// TIA Portal V20 export
Screen "CycleTime"  1276x673
  ScreenItem "Faceplate container_1" at 135,81 size 64x420  Type=HmiFaceplateContainer
  ScreenItem "Line_22" at 128,84 size 1x400  Type=HmiLine
  ScreenItem "Line_46" at 110,355 size 17x0  Type=HmiLine
  ScreenItem "Line_47" at 111,420 size 17x0  Type=HmiLine
  ScreenItem "Line_48" at 112,484 size 17x0  Type=HmiLine
  ScreenItem "Casella di testo_56" at 62,271 size 48x30  Type=HmiTextBox
  ScreenItem "Casella di testo_57" at 62,339 size 48x30  Type=HmiTextBox
  ScreenItem "Casella di testo_59" at 62,405 size 48x30  Type=HmiTextBox
  ScreenItem "Casella di testo_60" at 62,468 size 48x30  Type=HmiTextBox
  ScreenItem "Line_49" at 109,224 size 17x0  Type=HmiLine
  ScreenItem "Casella di testo_7" at 62,209 size 48x30  Type=HmiTextBox
  ScreenItem "Casella di testo_8" at 62,143 size 48x30  Type=HmiTextBox
  ScreenItem "Line_50" at 109,158 size 17x0  Type=HmiLine
  ScreenItem "Line_51" at 109,103 size 17x0  Type=HmiLine
  ScreenItem "Line_52" at 110,286 size 17x0  Type=HmiLine
  ScreenItem "Casella di testo_27" at 87,577 size 151x35  Type=HmiTextBox
  ScreenItem "Casella di testo_31" at 171,577 size 151x35  Type=HmiTextBox
  ScreenItem "Casella di testo_32" at 242,577 size 151x35  Type=HmiTextBox
  ScreenItem "Casella di testo_35" at 310,577 size 151x35  Type=HmiTextBox
  ScreenItem "Casella di testo_37" at 388,577 size 151x35  Type=HmiTextBox
  ScreenItem "Casella di testo_38" at 460,577 size 151x35  Type=HmiTextBox
  ScreenItem "Casella di testo_39" at 524,577 size 151x35  Type=HmiTextBox
  ScreenItem "Casella di testo_40" at 597,577 size 151x35  Type=HmiTextBox
  ScreenItem "Casella di testo_41" at 671,577 size 151x35  Type=HmiTextBox
  ScreenItem "Casella di testo_42" at 739,577 size 151x35  Type=HmiTextBox
  ScreenItem "Casella di testo_43" at 809,577 size 151x35  Type=HmiTextBox
  ScreenItem "Casella di testo_44" at 884,577 size 151x35  Type=HmiTextBox
  ScreenItem "Casella di testo_45" at 955,577 size 151x35  Type=HmiTextBox
  ScreenItem "Casella di testo_46" at 1026,577 size 151x35  Type=HmiTextBox
  ScreenItem "Casella di testo_47" at 1106,577 size 151x35  Type=HmiTextBox
  ScreenItem "Faceplate container_2" at 206,81 size 64x420  Type=HmiFaceplateContainer
  ScreenItem "Faceplate container_3" at 277,81 size 64x420  Type=HmiFaceplateContainer
  ScreenItem "Faceplate container_4" at 348,81 size 64x420  Type=HmiFaceplateContainer
  ScreenItem "Faceplate container_5" at 419,81 size 64x420  Type=HmiFaceplateContainer
  ScreenItem "Faceplate container_6" at 490,81 size 64x420  Type=HmiFaceplateContainer
  ScreenItem "Faceplate container_7" at 563,81 size 64x420  Type=HmiFaceplateContainer
  ScreenItem "Faceplate container_8" at 634,81 size 64x420  Type=HmiFaceplateContainer
  ScreenItem "Faceplate container_9" at 707,81 size 64x420  Type=HmiFaceplateContainer
  ScreenItem "Faceplate container_10" at 778,81 size 64x420  Type=HmiFaceplateContainer
  ScreenItem "Faceplate container_11" at 927,81 size 64x420  Type=HmiFaceplateContainer
  ScreenItem "Faceplate container_12" at 993,81 size 64x420  Type=HmiFaceplateContainer
  ScreenItem "Faceplate container_13" at 1066,81 size 64x420  Type=HmiFaceplateContainer
  ScreenItem "Faceplate container_14" at 850,81 size 64x420  Type=HmiFaceplateContainer
  ScreenItem "Faceplate container_15" at 1139,81 size 64x420  Type=HmiFaceplateContainer
  ScreenItem "Line_23" at 133,286 size 1103x1  Type=HmiLine
  ScreenItem "Line_45" at 130,483 size 1110x1  Type=HmiLine
  ScreenItem "Casella di testo_26" at 6,6 size 1267x47  Type=HmiTextBox
  ScreenItem "Move_Legend" at 1183,7 size 90x44  Type=HmiButton
  ScreenItem "Casella di testo_1" at -34,295 size 145x35  Type=HmiTextBox
  ScreenItem "Line_1" at 39,168 size 1x122  Type=HmiLine
  ScreenItem "Casella di testo_2" at 626,614 size 67x30  Type=HmiTextBox
  ScreenItem "Line_2" at 757,566 size 1x122  Type=HmiLine
